// TIA Portal V21 export
TextList "TL_ListSt"  ListRange=Decimal
  TextListEntry   Text="čeka"
  TextListEntry   From=1, To=1, Text="gotovo"
  TextListEntry   From=2, To=2, Text="preskočeno"
  TextListEntry   From=3, To=3, Text="u tijeku"
